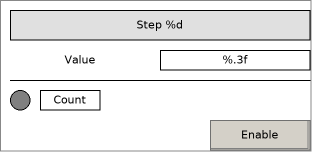
VISUALIZATION VISU_Fixture  // 312x152
    Rectangle (10,10 300x30), "Step %d", text variable: MAIN.fbStepChain.Step, colour toggle: GVL_Fixture.bEnable
    Label (10,50 140x20), "Value"
    Textfield (160,50 150x20), "%.3f", text variable: GVL_Fixture.fValue
    Line (10,80) (310,80)
    Ellipse (10,90 20x20), colour toggle: GVL_Fixture.bEnable
    RoundedRectangle (40,90 60x20), "Count", invisible if: NOT GVL_Fixture.bEnable
        p3560616238: GVL_Fixture.nCount
    Button (210,120 100x30), "Enable"
        p55702900: SEL(GVL_Fixture.bEnable, 16#FF000000, 16#FF00C000)
END_VISUALIZATION

(* stored: Version 1.1.0.1
   Visu VISU_Fixture: Id {4e4277b3-29d8-4ce6-9de1-2b0ca0bbbe8d} *)
